FUNCTION_BLOCK WaitMacro
VAR_INPUT
	Start 							: BOOL;
	WaitTime						: TIME;
END_VAR
VAR_OUTPUT
	Busy 							: BOOL;
	Done							: BOOL;
END_VAR
VAR
	state 							: UINT;
	fbStartTrigger					: R_TRIG;
	startTriggerOutput				: BOOL;
	fbTimerOn 						: TON;
	fbTimerOnStart					: BOOL;
	fbTimerOnEnd 					: BOOL;
END_VAR

fbTimerOn(IN:=fbTimerOnStart, PT := WaitTime, Q => fbTimerOnEnd);
fbStartTrigger(CLK := Start, Q => startTriggerOutput);
		
CASE state OF
	(************************** state 0 - IDLE *************************)  
	0:	
		Busy := FALSE;
		Done := FALSE;
		
		IF startTriggerOutput THEN
			Busy := TRUE;
			fbTimerOnStart := TRUE;
			state := 10;
		END_IF
	10:
		IF fbTimerOnEnd OR (WaitTime = T#0MS) THEN
			fbTimerOnStart := FALSE;
			state := 100;
		END_IF
	
	(************** state 100 - End *************)  
	100:
		Done := TRUE;
		state := 0;
		
END_CASE

END_FUNCTION_BLOCK

(* stored: Version 1.1.0.1, ProductVersion 3.1.4024.12
   POU WaitMacro: Id {48495372-d230-42ba-8dfc-c954e4f636c5}, SpecialFunc None *)
